FUNCTION_BLOCK FB_HeatPumpBuffer
VAR_INPUT
END_VAR
VAR_OUTPUT
	{attribute 'OPC.UA.DA' := '1'}	
	localState : ST_HeatPumpBufferState;
END_VAR
VAR
	MidTemperatureSensor : FB_TemperatureSensor_KL3214; //mid temperature sensor
END_VAR

//sensors
MidTemperatureSensor();

//get sensor inputs
MidTemperatureSensor.GetState_AI();

//set outputs
localState.fMidTemperature := MidTemperatureSensor.fTemperature;

END_FUNCTION_BLOCK

(* stored: Version 1.1.0.1
   POU FB_HeatPumpBuffer: Id {973783de-1af7-4dfe-b493-a43b76954c23}, SpecialFunc None *)
